Fanuc KAREL source: KT00660.KL

PROGRAM KT00660
%NOLOCKGROUP
VAR
  P1: POSITION
  P2: POSITION
  OUT: BOOLEAN
BEGIN
  OUT = - P1
END KT00660
